(* IEC 61131-3 sources: plc-hackathon-2026/evals/e3-compile-errors/src, 2 files *)

(* ---- E_Mode.st ---- *)
TYPE E_Mode :
(
    OFF := 0,
    AUTO,
    MANUAL
);
END_TYPE

(* ---- SR_Main.st ---- *)
PROGRAM SR_Main
VAR
    eMode  : E_Mode;
    iCount : INT;
    xOut   : BOOL;
END_VAR
// ---IMPL---
IF eMode = AUTO THEN
    iCount := iCount + 1
END_IF
xOut := iCount;
rTemp := 1.5;
